FUNCTION_BLOCK MoveArm (* Basic Function Block Type *)
  (* Standard: 61499-2 *)
  (* Version 0.0, 7/2/2026, Template *)
  PACKAGE Main;
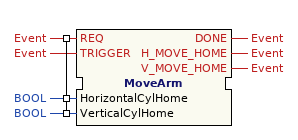
  EVENT_INPUT
    REQ WITH HorizontalCylHome, VerticalCylHome; (* Normal Execution Request *)
    TRIGGER; (* Initialization Request *)
  END_EVENT
  EVENT_OUTPUT
    DONE; (* Initialization Confirm *)
    H_MOVE_HOME; (* Execution Confirmation *)
    V_MOVE_HOME;
  END_EVENT
  VAR_INPUT
    HorizontalCylHome : BOOL; (* Input event qualifier *)
    VerticalCylHome : BOOL;
  END_VAR
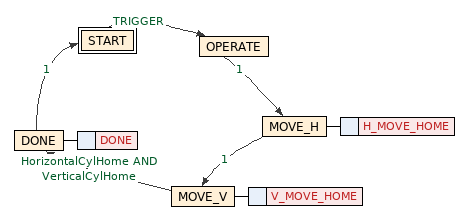
  EC_STATES
    START; (* Initial State *)
    OPERATE;
    MOVE_H : -> H_MOVE_HOME;
    MOVE_V : -> V_MOVE_HOME;
    DONE : -> DONE;
  END_STATES
  EC_TRANSITIONS
    START TO OPERATE := TRIGGER;
    OPERATE TO MOVE_H := 1;
    MOVE_H TO MOVE_V := 1;
    MOVE_V TO DONE := HorizontalCylHome AND VerticalCylHome;
    DONE TO START := 1;
  END_TRANSITIONS
  ALGORITHM INIT IN ST: (* Initialization algorithm *)
;
  END_ALGORITHM
  ALGORITHM REQ IN ST: (* Normally executed algorithm *)
;
  END_ALGORITHM
END_FUNCTION_BLOCK
